Yaskawa INFORM job: PICKDROP.JBI

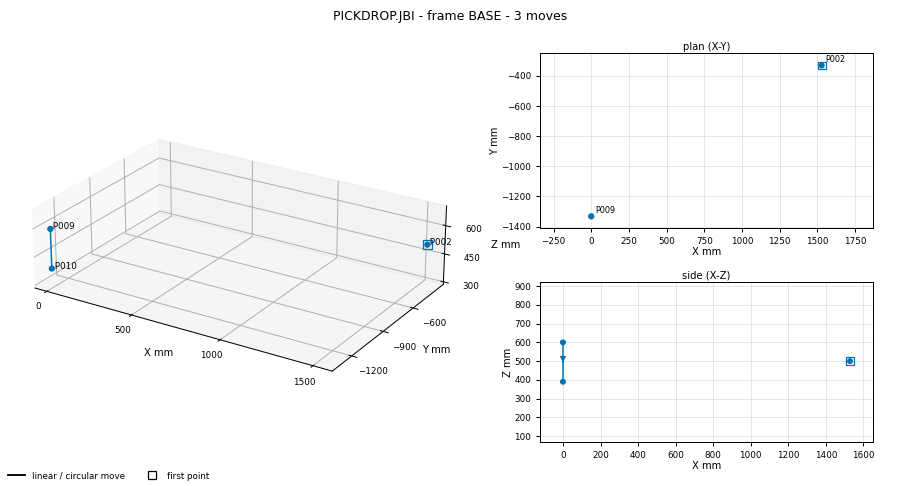
[picture p0: tool path of PICKDROP.JBI in frame BASE, 3 of 6 moves have a stored position in this frame; points joined in program order, loops and branches not executed]
/JOB
//NAME PICKDROP
//POS
///NPOS 0,0,0,6,0,0
///TOOL 0
///POSTYPE BASE
///RECTAN
///RCONF 1,0,0,0,1,0,0,0
P0002=1529.187,-331.251,500.000,180.00,0.00,90.00
///RCONF 0,0,0,0,0,0,0,0
P0003=0.000,0.000,-600.000,0.00,0.00,0.00
P0008=0.000,0.000,300.000,0.00,0.00,0.00
P0009=0.000,-1332.000,600.000,180.00,0.00,0.00
P0010=0.000,-1332.000,390.000,180.00,0.00,0.00
P0011=0.000,0.000,200.000,0.00,0.00,0.00
//INST
///DATE 2026/10/27 19:15
///ATTR SC,RW
///GROUP1 RB1
NOP
SET B090 0
SET B091 0
MOVL P002 V=I000 PL=0 DEC=50
IMOV P003 V=23.0 PL=0 BF UNTIL IN#(1)=ON
JUMP *FAULT IF IN#(1)=OFF
HAND HNO: 2 ON
SET I001 0
*CHECK
JUMP *VERIFY IF IN#(2)=ON
JUMP *VERIFY IF IN#(3)=ON
*VERIFY
TIMER T=0.10
INC I001
JUMP *FAULT IF I001>=10
JUMP *OK IF IN#(2)=ON
JUMP *OK IF IN#(3)=ON
JUMP *CHECK
*OK
IMOV P008 V=I000 PL=0 DEC=50
MOVL P009 V=I000 PL=0 DEC=50
SET B090 1
MOVL P010 V=I000 PL=0 DEC=50
HAND HNO: 2 OFF
TIMER T=1.00
IMOV P011 V=I000 PL=0
SET B091 1
JUMP *FINISH
*FAULT
SET B091 2
*HALT
PAUSE
JUMP *HALT
*FINISH
END
